(* IEC 61131-3 sources: IT-OT/examples, 5 files *)

(* ---- messwerte.st ---- *)
(* Messwerterfassung mit gleitendem Mittelwert.
   Zeigt: ARRAY, eigener FUNCTION_BLOCK, eigene FUNCTION.
   S7:     Rohwerte = DB1.DBW0 … DB1.DBW6 (4 Kanäle)
   OPC UA: ns=2;s=Rohwerte (Array), ns=2;s=Mittelwerte *)

FUNCTION Skaliere : REAL
VAR_INPUT
  Roh : INT;              (* 0 … 27648 wie bei S7-Analogeingängen *)
  Bereich : REAL := 100.0;
END_VAR
Skaliere := INT_TO_REAL(Roh) / 27648.0 * Bereich;
END_FUNCTION

FUNCTION_BLOCK GleitenderMittelwert
VAR_INPUT
  Wert : REAL;
END_VAR
VAR_OUTPUT
  Mittel : REAL;
  Gefuellt : BOOL;          (* Puffer einmal voll *)
END_VAR
VAR CONSTANT
  N : INT := 8;
END_VAR
VAR
  Puffer : ARRAY[0..7] OF REAL;
  Pos : INT;
  Summe : REAL;
  k : INT;
END_VAR
Puffer[Pos] := Wert;
Pos := (Pos + 1) MOD N;
IF Pos = 0 THEN Gefuellt := TRUE; END_IF;
Summe := 0.0;
FOR k := 0 TO N - 1 DO
  Summe := Summe + Puffer[k];
END_FOR;
Mittel := Summe / INT_TO_REAL(N);
END_FUNCTION_BLOCK

PROGRAM Messwerte
VAR_INPUT
  Rohwerte : ARRAY[0..3] OF INT := [13824, 27648, 0, 6912];
  Grenzwert : REAL := 80.0;
END_VAR
VAR_OUTPUT
  Mittelwerte : ARRAY[0..3] OF REAL;
  Alarm : ARRAY[0..3] OF BOOL;
  Bereit : BOOL;
END_VAR
VAR
  Filter0, Filter1, Filter2, Filter3 : GleitenderMittelwert;
  i : INT;
END_VAR
Filter0(Wert := Skaliere(Rohwerte[0]));
Filter1(Wert := Skaliere(Rohwerte[1]));
Filter2(Wert := Skaliere(Rohwerte[2]));
Filter3(Wert := Skaliere(Roh := Rohwerte[3], Bereich := 100.0));
Mittelwerte[0] := Filter0.Mittel;
Mittelwerte[1] := Filter1.Mittel;
Mittelwerte[2] := Filter2.Mittel;
Mittelwerte[3] := Filter3.Mittel;
FOR i := 0 TO 3 DO
  Alarm[i] := Mittelwerte[i] > Grenzwert;
END_FOR;
Bereit := Filter0.Gefuellt AND Filter1.Gefuellt AND Filter2.Gefuellt AND Filter3.Gefuellt;
END_PROGRAM

(* ---- ampel.st ---- *)
(* Fußgängerampel als Schrittkette.
   S7:     Anforderung = DB1.DBX0.0
   OPC UA: ns=2;s=Anforderung *)
PROGRAM Ampel
VAR CONSTANT
  T_GELB  : TIME := T#2s;
  T_ROT   : TIME := T#5s;
  T_RESET : TIME := T#1s;
END_VAR
VAR_INPUT
  Anforderung : BOOL;          (* Taster Fußgänger *)
END_VAR
VAR_OUTPUT
  Auto_Rot, Auto_Gelb, Auto_Gruen : BOOL;
  Fuss_Rot, Fuss_Gruen : BOOL;
  Zyklen : DINT;                (* Anzahl Fußgängerphasen *)
END_VAR
VAR
  Schritt : INT := 0;
  Timer   : TON;
  Taster  : R_TRIG;
  Angefordert : BOOL;
END_VAR

Taster(CLK := Anforderung);
IF Taster.Q THEN
  Angefordert := TRUE;
END_IF;

CASE Schritt OF
  0: (* Autos grün *)
     Auto_Gruen := TRUE; Auto_Gelb := FALSE; Auto_Rot := FALSE;
     Fuss_Rot := TRUE;  Fuss_Gruen := FALSE;
     IF Angefordert THEN
       Schritt := 10;
     END_IF;
  10: (* Autos gelb *)
     Auto_Gruen := FALSE; Auto_Gelb := TRUE;
     Timer(IN := TRUE, PT := T_GELB);
     IF Timer.Q THEN Timer(IN := FALSE); Schritt := 20; END_IF;
  20: (* Autos rot, Fußgänger grün *)
     Auto_Gelb := FALSE; Auto_Rot := TRUE;
     Fuss_Rot := FALSE; Fuss_Gruen := TRUE;
     Timer(IN := TRUE, PT := T_ROT);
     IF Timer.Q THEN Timer(IN := FALSE); Schritt := 30; END_IF;
  30: (* Räumzeit *)
     Fuss_Gruen := FALSE; Fuss_Rot := TRUE;
     Timer(IN := TRUE, PT := T_RESET);
     IF Timer.Q THEN
       Timer(IN := FALSE);
       Angefordert := FALSE;
       Zyklen := Zyklen + 1;
       Schritt := 0;
     END_IF;
ELSE
  Schritt := 0;
END_CASE;
END_PROGRAM

(* ---- foerderband.st ---- *)
(* Förderband mit Teilezählung, Losgröße und Störungsüberwachung. *)
PROGRAM Foerderband
VAR_INPUT
  Start, Stopp, Quittieren : BOOL;
  Sensor_Teil : BOOL;           (* Lichtschranke *)
  Losgroesse  : INT := 10;
END_VAR
VAR_OUTPUT
  Motor   : BOOL;
  Los_Fertig, Stoerung : BOOL;
  Teile   : INT;
  Gesamt  : UDINT;
END_VAR
VAR
  Zaehler : CTU;
  Teil    : R_TRIG;
  Laufzeit_Ohne_Teil : TON;
  Ein     : SR;
END_VAR

Ein(S1 := Start AND NOT Stoerung, R := Stopp OR Stoerung OR Los_Fertig);
Motor := Ein.Q1;

Teil(CLK := Sensor_Teil);
IF Teil.Q THEN Gesamt := Gesamt + 1; END_IF;

Zaehler(CU := Teil.Q, R := Quittieren, PV := Losgroesse);
Teile := Zaehler.CV;
Los_Fertig := Zaehler.Q;

(* Störung: Band läuft 10 s ohne dass ein Teil erkannt wird *)
Laufzeit_Ohne_Teil(IN := Motor AND NOT Sensor_Teil, PT := T#10s);
IF Laufzeit_Ohne_Teil.Q THEN
  Stoerung := TRUE;
END_IF;
IF Quittieren THEN
  Stoerung := FALSE;
END_IF;
END_PROGRAM

(* ---- lager.st ---- *)
(* Kleines Lager mit 5 Fächern.
   Zeigt: TYPE … STRUCT (UDT), Arrays von Strukturen, STRING und String-Funktionen.
   Einlagern: Artikel, Menge und Fach setzen, dann Buchen auf TRUE.
   OPC UA: ns=2;s=Faecher[2].Artikel, ns=2;s=Meldung
   API:    PUT /api/plcs/Lager/variables/Auftrag  {"value": {"Artikel": "Schraube M6", "Menge": 50, "Fach": 2}} *)

TYPE
  Lagerfach : STRUCT
    Artikel : STRING[20];
    Menge   : INT;
    Gesperrt : BOOL;
  END_STRUCT;
  Buchung : STRUCT
    Artikel : STRING[20];
    Menge   : INT;      (* positiv = einlagern, negativ = auslagern *)
    Fach    : INT := 1;
  END_STRUCT;
END_TYPE

PROGRAM Lager
VAR_INPUT
  Auftrag : Buchung;
  Buchen  : BOOL;
END_VAR
VAR_OUTPUT
  Faecher : ARRAY[1..5] OF Lagerfach;
  Bestand : DINT;
  Meldung : STRING[60] := 'Bereit';
  Fehler  : BOOL;
END_VAR
VAR
  Flanke : R_TRIG;
  i : INT;
END_VAR

Flanke(CLK := Buchen);
IF Flanke.Q THEN
  Fehler := TRUE;
  IF Auftrag.Fach < 1 OR Auftrag.Fach > 5 THEN
    Meldung := CONCAT('Fach ungültig: ', INT_TO_STRING(Auftrag.Fach));
  ELSIF Faecher[Auftrag.Fach].Gesperrt THEN
    Meldung := CONCAT('Fach gesperrt: ', INT_TO_STRING(Auftrag.Fach));
  ELSIF Faecher[Auftrag.Fach].Menge > 0 AND Faecher[Auftrag.Fach].Artikel <> Auftrag.Artikel THEN
    Meldung := CONCAT('Fach belegt mit ', Faecher[Auftrag.Fach].Artikel);
  ELSIF Faecher[Auftrag.Fach].Menge + Auftrag.Menge < 0 THEN
    Meldung := 'Zu wenig Bestand';
  ELSE
    Faecher[Auftrag.Fach].Artikel := Auftrag.Artikel;
    Faecher[Auftrag.Fach].Menge := Faecher[Auftrag.Fach].Menge + Auftrag.Menge;
    IF Faecher[Auftrag.Fach].Menge = 0 THEN
      Faecher[Auftrag.Fach].Artikel := '';
    END_IF;
    Meldung := CONCAT(CONCAT(INT_TO_STRING(Auftrag.Menge), ' x '), Auftrag.Artikel);
    Fehler := FALSE;
  END_IF;
END_IF;

Bestand := 0;
FOR i := 1 TO 5 DO
  Bestand := Bestand + Faecher[i].Menge;
END_FOR;
END_PROGRAM

(* ---- tank.st ---- *)
(* Füllstandsregelung mit Zweipunktregler und simulierter Strecke.
   Ideal zum Testen von HMI/SCADA-Anbindungen über S7 oder OPC UA. *)
PROGRAM Tank
VAR_INPUT
  Automatik : BOOL := TRUE;
  Sollwert  : REAL := 60.0;    (* % *)
  Hysterese : REAL := 5.0;     (* % *)
  Abfluss   : REAL := 0.15;    (* %/Zyklus *)
END_VAR
VAR_OUTPUT
  Fuellstand : REAL := 20.0;   (* % *)
  Pumpe      : BOOL;
  Alarm_Hoch, Alarm_Tief : BOOL;
  Pumpenstarts : DINT;
END_VAR
VAR
  Zufluss : REAL := 0.4;
  Start   : R_TRIG;
  Alarm_Verz : TON;
END_VAR

IF Automatik THEN
  IF Fuellstand < Sollwert - Hysterese THEN
    Pumpe := TRUE;
  ELSIF Fuellstand > Sollwert + Hysterese THEN
    Pumpe := FALSE;
  END_IF;
END_IF;

Start(CLK := Pumpe);
IF Start.Q THEN Pumpenstarts := Pumpenstarts + 1; END_IF;

(* Simulation der Strecke *)
IF Pumpe THEN
  Fuellstand := Fuellstand + Zufluss;
END_IF;
Fuellstand := LIMIT(0.0, Fuellstand - Abfluss, 100.0);

Alarm_Verz(IN := Fuellstand > 95.0 OR Fuellstand < 5.0, PT := T#2s);
Alarm_Hoch := Alarm_Verz.Q AND Fuellstand > 95.0;
Alarm_Tief := Alarm_Verz.Q AND Fuellstand < 5.0;
END_PROGRAM
